# EPICS autosave request: iocs/meascomp/db/measCompWaveformGen_settings.req
$(P)$(R)UserNumPoints
$(P)$(R)IntNumPoints
$(P)$(R)UserDwell
$(P)$(R)IntDwell
$(P)$(R)ExtTrigger
$(P)$(R)ExtClock
$(P)$(R)Continuous
$(P)$(R)Retrigger
$(P)$(R)TriggerCount
